// TIA Portal V20 export
FUNCTION_BLOCK "FB_BatchSequence"   // FB104, GRAPH
TITLE = Batch sequence: fill A, fill B, mix and heat, hold, drain
AUTHOR : Demo
VERSION : 0.2
// GRAPH version. Same inputs and outputs as scl/16_FB_BatchSequence.scl.
// stored: GraphVersion 2.0, SetENOAutomatically false
   // inherited from GRAPH_BASE
   VAR_INPUT
      OFF_SQ : Bool;
      INIT_SQ : Bool;
      ACK_EF : Bool;
      S_PREV : Bool;
      S_NEXT : Bool;
      SW_AUTO : Bool;
      SW_TAP : Bool;
      SW_TOP : Bool;
      SW_MAN : Bool;
      S_SEL : Int;
      S_ON : Bool;
      S_OFF : Bool;
      T_PUSH : Bool;
      Start : Bool;   // Start button or MES start request
      Stop : Bool;   // Stop button: pause the batch
      Auto : Bool;   // Selector in Auto
      AnyFault : Bool;   // Any FAULT alarm active
      EStopOK : Bool;   // Emergency stop circuit healthy
      Level : Real;   // Tank level [%]
      Temp : Real;   // Tank temperature [degC]
      FillerReady : Bool;   // Downstream filler ready to receive
   END_VAR
   VAR_OUTPUT
      S_NO : Int;
      S_MORE : Bool;
      S_ACTIVE : Bool;
      ERR_FLT : Bool;
      AUTO_ON : Bool;
      TAP_ON : Bool;
      TOP_ON : Bool;
      MAN_ON : Bool;
      "Step" : Int;   // Current step: 0 Idle, 10 Fill A, 20 Fill B, 30 Mix and heat, 40 Hold, 50 Drain, 60 Done
      StepTime : Time;   // Time in the current step without interlock error (pauses while halted)
      Halted : Bool;   // Sequence paused: outputs off (fault, E-stop, Stop or not in Auto)
      Running : Bool;   // A batch is active (step 10..60)
      OpenXV101 : Bool;   // Command: open inlet valve A
      OpenXV102 : Bool;   // Command: open inlet valve B
      RunM201 : Bool;   // Command: run agitator
      SpeedM201 : Real;   // Command: agitator speed [rpm]
      HeatE301 : Bool;   // Command: heater on
      RunP401 : Bool;   // Command: run outlet pump
      BatchDone : Bool;   // Pulse when a batch finishes
      RecipeValid : Bool;   // Recipe values are plausible
      TimeoutStep10 : Bool;   // Step 10 longer than 120 s
      TimeoutStep20 : Bool;   // Step 20 longer than 120 s
      TimeoutStep30 : Bool;   // Step 30 longer than 600 s
      TimeoutStep50 : Bool;   // Step 50 longer than 180 s
      WaitFillerTooLong : Bool;   // Step 40 waiting for filler longer than 60 s
      StartNotAuto : Bool;   // Start pressed while not in Auto
      StartTankNotEmpty : Bool;   // Start pressed while tank not empty
      StartRecipeInvalid : Bool;   // Start pressed while recipe invalid
   END_VAR
   VAR
      Paused : Bool;   // Set by Stop, a fault or the E-stop; cleared by Start
      Healthy : Bool;   // No fault, E-stop OK, not paused and in Auto: the step interlocks are fulfilled
      HeatReq : Bool;   // Step 30 asks for heat (heater runs while below TempSP)
   END_VAR
BEGIN
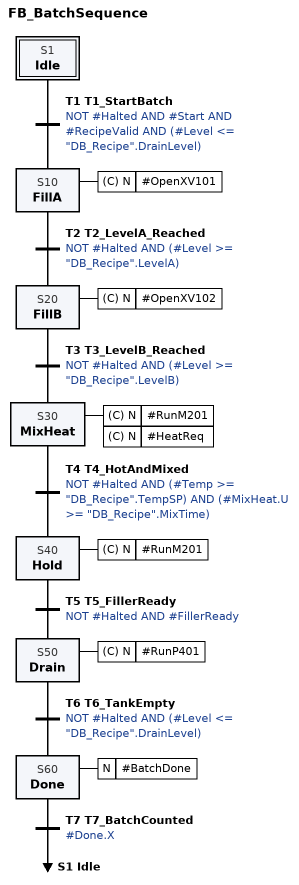
   // permanent pre-instructions
   NETWORK 1
      #RecipeValid := ("DB_Recipe".LevelA > 0.0) AND ("DB_Recipe".LevelA < "DB_Recipe".LevelB) AND ("DB_Recipe".LevelB <= 90.0) AND ("DB_Recipe".TempSP >= 20.0) AND ("DB_Recipe".TempSP <= 85.0) AND ("DB_Recipe".MixSpeed >= 100.0) AND ("DB_Recipe".MixSpeed <= 1500.0);
   NETWORK 2
      IF #Start THEN #Paused := FALSE; END_IF;
   NETWORK 3
      IF #Stop THEN #Paused := TRUE; END_IF;
   NETWORK 4
      IF #AnyFault THEN #Paused := TRUE; END_IF;
   NETWORK 5
      IF NOT #EStopOK THEN #Paused := TRUE; END_IF;
   NETWORK 6
      #Healthy := NOT #AnyFault AND #EStopOK AND NOT #Paused AND #Auto;
   NETWORK 7
      #Halted := NOT #Healthy;

   // sequencer 1
   // Batch sequence of the mixing station. Idle waits for Start; Fill A and Fill B open the inlet valves until the recipe levels; Mix and heat runs the agitator and heats to TempSP for MixTime; Hold waits for the filler; Drain pumps the tank empty; Done counts the batch. Every working step is interlocked with Healthy: on a fault, E-stop, Stop or Auto off its actions switch off and the step is kept. After a fault or E-stop, press Reset, then Start to continue; Reset alone does not restart the batch.
   INITIAL_STEP Idle:   // S1, max time T#10S, warning time T#10S
   END_STEP
   TRANSITION T1_StartBatch FROM Idle TO FillA   // T1
      := NOT #Halted AND #Start AND #RecipeValid AND (#Level <= "DB_Recipe".DrainLevel);
   END_TRANSITION
   STEP FillA:   // S10, max time T#120S, warning time T#120S
      interlock C := #Healthy;   // Sequence halted: fault, E-stop, Stop or not in Auto
      (C)     N    #OpenXV101
   END_STEP
   TRANSITION T2_LevelA_Reached FROM FillA TO FillB   // T2
      := NOT #Halted AND (#Level >= "DB_Recipe".LevelA);
   END_TRANSITION
   STEP FillB:   // S20, max time T#120S, warning time T#120S
      interlock C := #Healthy;   // Sequence halted: fault, E-stop, Stop or not in Auto
      (C)     N    #OpenXV102
   END_STEP
   TRANSITION T3_LevelB_Reached FROM FillB TO MixHeat   // T3
      := NOT #Halted AND (#Level >= "DB_Recipe".LevelB);
   END_TRANSITION
   STEP MixHeat:   // S30, max time T#600S, warning time T#600S
      interlock C := #Healthy;   // Sequence halted: fault, E-stop, Stop or not in Auto
      (C)     N    #RunM201
      (C)     N    #HeatReq
   END_STEP
   TRANSITION T4_HotAndMixed FROM MixHeat TO Hold   // T4
      := NOT #Halted AND (#Temp >= "DB_Recipe".TempSP) AND (#MixHeat.U >= "DB_Recipe".MixTime);
   END_TRANSITION
   STEP Hold:   // S40, max time T#60S, warning time T#60S
      interlock C := #Healthy;   // Sequence halted: fault, E-stop, Stop or not in Auto
      (C)     N    #RunM201
   END_STEP
   TRANSITION T5_FillerReady FROM Hold TO Drain   // T5
      := NOT #Halted AND #FillerReady;
   END_TRANSITION
   STEP Drain:   // S50, max time T#180S, warning time T#180S
      interlock C := #Healthy;   // Sequence halted: fault, E-stop, Stop or not in Auto
      (C)     N    #RunP401
   END_STEP
   TRANSITION T6_TankEmpty FROM Drain TO Done   // T6
      := NOT #Halted AND (#Level <= "DB_Recipe".DrainLevel);
   END_TRANSITION
   STEP Done:   // S60, max time T#10S, warning time T#10S
              N    #BatchDone
   END_STEP
   TRANSITION T7_BatchCounted FROM Done TO Idle   // T7, jump
      := #Done.X;
   END_TRANSITION

   // permanent post-instructions
   NETWORK 1
      IF #Idle.X THEN
          #"Step" := 0;
          #StepTime := #Idle.U;
      END_IF;
   NETWORK 2
      IF #FillA.X THEN
          #"Step" := 10;
          #StepTime := #FillA.U;
      END_IF;
   NETWORK 3
      IF #FillB.X THEN
          #"Step" := 20;
          #StepTime := #FillB.U;
      END_IF;
   NETWORK 4
      IF #MixHeat.X THEN
          #"Step" := 30;
          #StepTime := #MixHeat.U;
      END_IF;
   NETWORK 5
      IF #Hold.X THEN
          #"Step" := 40;
          #StepTime := #Hold.U;
      END_IF;
   NETWORK 6
      IF #Drain.X THEN
          #"Step" := 50;
          #StepTime := #Drain.U;
      END_IF;
   NETWORK 7
      IF #Done.X THEN
          #"Step" := 60;
          #StepTime := #Done.U;
      END_IF;
   NETWORK 8
      #Running := NOT #Idle.X;
   NETWORK 9
      IF #MixHeat.X THEN #SpeedM201 := "DB_Recipe".MixSpeed; END_IF;
   NETWORK 10
      IF NOT #MixHeat.X THEN #SpeedM201 := "DB_Recipe".HoldSpeed; END_IF;
   NETWORK 11
      #HeatE301 := #HeatReq AND (#Temp < "DB_Recipe".TempSP);
   NETWORK 12
      #TimeoutStep10 := #FillA.X AND (#FillA.U > T#120S);
   NETWORK 13
      #TimeoutStep20 := #FillB.X AND (#FillB.U > T#120S);
   NETWORK 14
      #TimeoutStep30 := #MixHeat.X AND (#MixHeat.U > T#600S);
   NETWORK 15
      #TimeoutStep50 := #Drain.X AND (#Drain.U > T#180S);
   NETWORK 16
      #WaitFillerTooLong := #Hold.X AND (#Hold.U > T#60S) AND NOT #FillerReady;
   NETWORK 17
      #StartNotAuto := #Idle.X AND #Start AND NOT #Auto;
   NETWORK 18
      #StartTankNotEmpty := #Idle.X AND #Start AND (#Level > "DB_Recipe".DrainLevel);
   NETWORK 19
      #StartRecipeInvalid := #Idle.X AND #Start AND NOT #RecipeValid;
END_FUNCTION_BLOCK
